// TIA Portal V19 export
DATA_BLOCK "Tacho2_EM05"   // DB6
VERSION : 1.0
// stored: InstanceOfName EM05_Agitacion, InstanceOfType FB
"EM05_Agitacion"
   // VAR_INPUT
   //    In : "EM05_Input";
   //    MotorFbkRun : Bool;
   //    MotorTrip : Bool;
   // END_VAR
   // VAR_OUTPUT
   //    Out : "EM05_Output";
   //    CM_Mot_Agitador_Out : Bool;
   //    CMAlarm : Bool;
   // END_VAR
   // VAR
   //    State : Int;
   //    ActiveAgitatorType : Int;
   //    AlarmLatched : Bool;
   //    FaultCode : Int;
   //    TrigStart { S7_SetPoint := 'True'} : R_TRIG;
   //    TrigStop { S7_SetPoint := 'True'} : R_TRIG;
   //    TrigHold { S7_SetPoint := 'True'} : R_TRIG;
   //    TrigAbort { S7_SetPoint := 'True'} : R_TRIG;
   //    TrigReset { S7_SetPoint := 'True'} : R_TRIG;
   //    CM_Mot_Agitador { S7_SetPoint := 'True'} : "MotL";
   // END_VAR
BEGIN
END_DATA_BLOCK
